DATA_BLOCK "naut_SfcJumpBack_DB"
{ S7_Optimized_Access := 'TRUE' }
VERSION : 0.1
"naut_SfcJumpBack"

BEGIN

END_DATA_BLOCK
